(* IEC 61131-3 sources: codesys-to-s7/tests/corpus/C2S7-LIB/pos, 1 file *)

(* ---- input.st ---- *)
FUNCTION_BLOCK FB_Case
VAR
    n : INT;
    a : INT;
END_VAR
n := SIZEOF(a);
END_FUNCTION_BLOCK
